(*
SPDX-FileCopyrightText: © 2026 Oleksandr Tiutyk <trofimich@gmail.com>
SPDX-License-Identifier: MIT
License: https://opensource.org/license/mit
*)

(*!
<summary>Checks safe defaults for an unbound TaskState view.</summary>
<description>
Uses unbound local references and checks every observable property without dereferencing a missing target.
</description>
*)

{attribute 'no_explicit_call' := 'do not call this function block directly'}
FUNCTION_BLOCK UnboundTaskStateTest EXTENDS TOF_Testing.SingleCycleTest
VAR_STAT
	{attribute 'hide'}
	_ClassName : STRING := __POUNAME();
END_VAR

//! <summary>Reads all flags and verifies the default value for an unbound view.</summary>
METHOD PROTECTED ExecuteTest
VAR
	backingValue : REFERENCE TO TOF_Tasks.TASK_STATE;
	stateChanged : REFERENCE TO BOOL;
	view : TOF_Tasks.TaskState(taskState := backingValue, taskStateChanged := stateChanged);
END_VAR
Assert.ThatBool(actual := view.Ready, message := "Unbound TaskState.Ready must be false").IsFalse();
Assert.ThatBool(actual := view.Running, message := "Unbound TaskState.Running must be false").IsFalse();
Assert.ThatBool(actual := view.Stopped, message := "Unbound TaskState.Stopped must be false").IsFalse();
Assert.ThatBool(actual := view.StateChanged, message := "Unbound TaskState.StateChanged must be false").IsFalse();
Assert.ThatBool(
	actual := view.Value = TOF_Tasks.TASK_STATE.READY,
	message := "Unbound Value must default to READY"
).IsTrue();
END_METHOD

//! <summary>Borrows the concrete class name. Callers must not modify the returned storage.</summary>
{attribute 'monitoring' := 'call'}
PROPERTY ClassName : REFERENCE TO STRING
GET
ClassName REF= _ClassName;
END_GET
END_PROPERTY

//! <summary>Borrows the compiler-initialized namespace name. Callers must not modify the returned storage.</summary>
{attribute 'monitoring' := 'call'}
PROPERTY NamespaceName : REFERENCE TO STRING
GET
NamespaceName REF= CurrentNamespace.Name;
END_GET
END_PROPERTY

//! <summary>Reports the complete concrete instance size in bytes.</summary>
{attribute 'monitoring' := 'call'}
PROPERTY SelfSize : ULINT
GET
SelfSize := XSIZEOF(THIS^);
END_GET
END_PROPERTY

END_FUNCTION_BLOCK

(* stored: Version 1.1.0.1
   POU UnboundTaskStateTest: Id {5c667417-1b52-4dd6-a1b8-23ce4dc6d4bc}, SpecialFunc None
   Method ExecuteTest: Id {a14d76e2-7fcd-4359-b9eb-0b80e7b5180e}
   Property ClassName: Id {29b14cf5-0836-447c-8c9e-c229ab6dee50}
   Get Get: Id {de7c0e28-26fe-47f5-b82e-b84da826e169}
   Property NamespaceName: Id {07370dcc-7f9b-4df2-ac23-6112ffe3bc23}
   Get Get: Id {aad4619a-78fb-46f6-ac18-17ef847dda45}
   Property SelfSize: Id {7d81fc7d-4ee3-445f-9688-ff05699259b7}
   Get Get: Id {1e0116ac-5fc6-435d-bab4-72e8defee532} *)
